METHOD PRIVATE Teach_OutOfTolerance_IsRejected
VAR_INST
    bRan : BOOL;
END_VAR
VAR
    stPlace : ST_SlotAddr := (nSide := 1, nColumn := 3, nLevel := 2);
END_VAR
TEST('Teach_OutOfTolerance_IsRejected');
IF bRan THEN
    TEST_FINISHED();
    RETURN;
END_IF
bRan := TRUE;

AssertFalse(Condition := fbRackReject.Teach(stPlace, fbRackReject.NominalX(stPlace) + 0.035, fbRackReject.NominalY(stPlace)),
            Message := '35 mm off the drawing means check the rack, not learn it');
AssertEquals_LREAL(Expected := fbRackReject.NominalX(stPlace), Actual := fbRackReject.TargetX(stPlace), Delta := 1.0E-9,
                   Message := 'a rejected teach must not change the target');

TEST_FINISHED();
END_METHOD

METHOD PRIVATE PutTake_BooksThePalletInAndOut
VAR_INST
    bRan : BOOL;
END_VAR
VAR
    stPlace : ST_SlotAddr := (nSide := 1, nColumn := 1, nLevel := 1);
END_VAR
TEST('PutTake_BooksThePalletInAndOut');
IF bRan THEN
    TEST_FINISHED();
    RETURN;
END_IF
bRan := TRUE;

AssertTrue(Condition := fbRackBook.Put(stPlace, 'LE0001'), Message := 'empty place must accept a pallet');
AssertTrue(Condition := fbRackBook.IsOccupied(stPlace), Message := 'place must be occupied after Put');
AssertEquals_STRING(Expected := 'LE0001', Actual := fbRackBook.LeIdAt(stPlace), Message := 'place must know its load unit');
AssertEquals_STRING(Expected := 'LE0001', Actual := fbRackBook.Take(stPlace), Message := 'Take must return the load unit');
AssertFalse(Condition := fbRackBook.IsOccupied(stPlace), Message := 'place must be free after Take');

TEST_FINISHED();
END_METHOD

METHOD PRIVATE Put_OnOccupiedPlace_IsRefused
VAR_INST
    bRan : BOOL;
END_VAR
VAR
    stPlace : ST_SlotAddr := (nSide := 2, nColumn := 7, nLevel := 4);
END_VAR
TEST('Put_OnOccupiedPlace_IsRefused');
IF bRan THEN
    TEST_FINISHED();
    RETURN;
END_IF
bRan := TRUE;

fbRackTwice.Put(stPlace, 'LE0001');
AssertFalse(Condition := fbRackTwice.Put(stPlace, 'LE0002'), Message := 'two pallets must never be booked into one place');
AssertEquals_STRING(Expected := 'LE0001', Actual := fbRackTwice.LeIdAt(stPlace), Message := 'first pallet must stay booked');

TEST_FINISHED();
END_METHOD

METHOD PRIVATE InvalidAddress_IsRejectedEverywhere
VAR_INST
    bRan : BOOL;
END_VAR
VAR
    stSide3 : ST_SlotAddr := (nSide := 3, nColumn := 1, nLevel := 1);
    stCol21 : ST_SlotAddr := (nSide := 1, nColumn := 21, nLevel := 1);
    stStationLevel2 : ST_SlotAddr := (nSide := 1, nColumn := 0, nLevel := 2);
END_VAR
TEST('InvalidAddress_IsRejectedEverywhere');
IF bRan THEN
    TEST_FINISHED();
    RETURN;
END_IF
bRan := TRUE;

AssertFalse(Condition := fbRackBad.IsValid(stSide3), Message := 'side 3 does not exist');
AssertFalse(Condition := fbRackBad.IsValid(stCol21), Message := 'column 21 does not exist');
AssertFalse(Condition := fbRackBad.IsValid(stStationLevel2), Message := 'the station has only level 1');
AssertFalse(Condition := fbRackBad.Put(stCol21, 'LE0001'), Message := 'no booking into an invalid address');

TEST_FINISHED();
END_METHOD

METHOD PRIVATE FindFree_SkipsOccupiedPlaces
VAR_INST
    bRan : BOOL;
END_VAR
VAR
    stA : ST_SlotAddr := (nSide := 1, nColumn := 1, nLevel := 1);
    stB : ST_SlotAddr := (nSide := 2, nColumn := 1, nLevel := 1);
    stFound : ST_SlotAddr;
END_VAR
TEST('FindFree_SkipsOccupiedPlaces');
IF bRan THEN
    TEST_FINISHED();
    RETURN;
END_IF
bRan := TRUE;

fbRackFree.Put(stA, 'LE0001');
fbRackFree.Put(stB, 'LE0002');
AssertTrue(Condition := fbRackFree.FindFree(stFound), Message := 'an almost empty rack has free places');
AssertEquals_INT(Expected := 1, Actual := stFound.nColumn, Message := 'nearest column first');
AssertEquals_INT(Expected := 2, Actual := stFound.nLevel, Message := 'level 1 is full on both sides -> level 2');

TEST_FINISHED();
END_METHOD

END_FUNCTION_BLOCK

// ---- Test/FB_Axis_Test.TcPOU
// Tests for FB_Axis, the simulated positioning axis. Each test drives the axis
// to the end inside one PLC cycle (simulated time), so they are fast.
FUNCTION_BLOCK FB_Axis_Test EXTENDS TcUnit.FB_TestSuite
VAR
    fbAxArrive  : FB_Axis(ipParent := 0, sNodeName := 'AxArrive');
    fbAxLong    : FB_Axis(ipParent := 0, sNodeName := 'AxLong');
    fbAxShort   : FB_Axis(ipParent := 0, sNodeName := 'AxShort');
    fbAxFault   : FB_Axis(ipParent := 0, sNodeName := 'AxFault');
    fbAxReset   : FB_Axis(ipParent := 0, sNodeName := 'AxReset');
END_VAR

Move_ArrivesInsideTheTolerance();
LongMove_TakesTheTrapezoidTime();
ShortMove_TakesTheTriangleTime();
DriveFault_WhileMoving_FailsTheMove();
Reset_AfterFault_AllowsTheNextMove();

METHOD PRIVATE Move_ArrivesInsideTheTolerance
VAR_INST
    bRan : BOOL;
END_VAR
VAR
    eResult : E_CmdResult;
    n : DINT;
END_VAR
TEST('Move_ArrivesInsideTheTolerance');
IF bRan THEN
    TEST_FINISHED();
    RETURN;
END_IF
bRan := TRUE;

FOR n := 1 TO 20000 DO
    eResult := fbAxArrive.MoveAbs(10.0);
    IF eResult <> E_CmdResult.eBusy THEN EXIT; END_IF
    fbAxArrive.Cyclic();
END_FOR
AssertTrue(Condition := eResult = E_CmdResult.eDone, Message := 'move must finish with eDone');
AssertEquals_LREAL(Expected := 10.0, Actual := fbAxArrive.lrActPos, Delta := fbAxArrive.lrTolerance, Message := 'axis must stand inside the tolerance');
AssertEquals_LREAL(Expected := 0.0, Actual := fbAxArrive.lrActVelo, Delta := 1.0E-9, Message := 'axis must stand still');

TEST_FINISHED();
END_METHOD

METHOD PRIVATE LongMove_TakesTheTrapezoidTime
VAR_INST
    bRan : BOOL;
END_VAR
VAR
    eResult : E_CmdResult;
    n : DINT;
    lrTime : LREAL;
END_VAR
TEST('LongMove_TakesTheTrapezoidTime');
IF bRan THEN
    TEST_FINISHED();
    RETURN;
END_IF
bRan := TRUE;

fbAxLong.lrVelocity := 3.0;
fbAxLong.lrAccel    := 0.6;
FOR n := 1 TO 20000 DO
    eResult := fbAxLong.MoveAbs(20.0);
    IF eResult <> E_CmdResult.eBusy THEN EXIT; END_IF
    fbAxLong.Cyclic();
    lrTime := lrTime + fbAxLong.lrCycleTime;
END_FOR
// 20 m >= v^2/a = 15 m -> top speed reached: t = s/v + v/a = 6.67 + 5.0 s
AssertEquals_LREAL(Expected := F_TravelTime(20.0, 3.0, 0.6), Actual := lrTime, Delta := 0.1, Message := 'move time must match s/v + v/a');

TEST_FINISHED();
END_METHOD

METHOD PRIVATE ShortMove_TakesTheTriangleTime
VAR_INST
    bRan : BOOL;
END_VAR
VAR
    eResult : E_CmdResult;
    n : DINT;
    lrTime : LREAL;
END_VAR
TEST('ShortMove_TakesTheTriangleTime');
IF bRan THEN
    TEST_FINISHED();
    RETURN;
END_IF
bRan := TRUE;

fbAxShort.lrVelocity := 3.0;
fbAxShort.lrAccel    := 0.6;
FOR n := 1 TO 20000 DO
    eResult := fbAxShort.MoveAbs(1.0);
    IF eResult <> E_CmdResult.eBusy THEN EXIT; END_IF
    fbAxShort.Cyclic();
    lrTime := lrTime + fbAxShort.lrCycleTime;
END_FOR
// 1 m < 15 m -> never reaches 3 m/s: t = 2 * sqrt(s/a) = 2.58 s
AssertEquals_LREAL(Expected := F_TravelTime(1.0, 3.0, 0.6), Actual := lrTime, Delta := 0.1, Message := 'short move must follow the triangle profile');

TEST_FINISHED();
END_METHOD

METHOD PRIVATE DriveFault_WhileMoving_FailsTheMove
VAR_INST
    bRan : BOOL;
END_VAR
VAR
    eResult : E_CmdResult;
    n : DINT;
END_VAR
TEST('DriveFault_WhileMoving_FailsTheMove');
IF bRan THEN
    TEST_FINISHED();
    RETURN;
END_IF
bRan := TRUE;

FOR n := 1 TO 50 DO
    fbAxFault.MoveAbs(5.0);
    fbAxFault.Cyclic();
END_FOR
fbAxFault.bDriveFault := TRUE;
fbAxFault.Cyclic();
eResult := fbAxFault.MoveAbs(5.0);
AssertTrue(Condition := eResult = E_CmdResult.eError, Message := 'a drive fault during a move must give eError');
AssertEquals_LREAL(Expected := 0.0, Actual := fbAxFault.lrActVelo, Delta := 1.0E-9, Message := 'a faulted axis must stand still');

TEST_FINISHED();
END_METHOD

METHOD PRIVATE Reset_AfterFault_AllowsTheNextMove
VAR_INST
    bRan : BOOL;
END_VAR
VAR
    eResult : E_CmdResult;
    n : DINT;
END_VAR
TEST('Reset_AfterFault_AllowsTheNextMove');
IF bRan THEN
    TEST_FINISHED();
    RETURN;
END_IF
bRan := TRUE;

fbAxReset.MoveAbs(5.0);
fbAxReset.Cyclic();
fbAxReset.bDriveFault := TRUE;
fbAxReset.Cyclic();
fbAxReset.bDriveFault := FALSE;
fbAxReset.Reset();
FOR n := 1 TO 20000 DO
    eResult := fbAxReset.MoveAbs(2.0);
    IF eResult <> E_CmdResult.eBusy THEN EXIT; END_IF
    fbAxReset.Cyclic();
END_FOR
AssertTrue(Condition := eResult = E_CmdResult.eDone, Message := 'after Reset a new move must work');

TEST_FINISHED();
END_METHOD

END_FUNCTION_BLOCK

// ---- Performance/F_TravelTime.TcPOU
// Time for one axis to travel lrDist with a trapezoid profile [s]:
// reaches top speed if lrDist >= v^2/a, otherwise a triangle profile.
FUNCTION F_TravelTime : LREAL
VAR_INPUT
    lrDist  : LREAL;   // [m]
    lrVelo  : LREAL;   // max. speed [m/s]
    lrAccel : LREAL;   // acceleration = deceleration [m/s2]
END_VAR
VAR
    lrD : LREAL;
END_VAR

lrD := ABS(lrDist);
IF lrD <= 0.0 OR lrVelo <= 0.0 OR lrAccel <= 0.0 THEN
    F_TravelTime := 0.0;
ELSIF lrD >= lrVelo * lrVelo / lrAccel THEN
    F_TravelTime := lrD / lrVelo + lrVelo / lrAccel;
ELSE
    F_TravelTime := 2.0 * SQRT(lrD / lrAccel);
END_IF

END_FUNCTION

// ---- Test/FB_ConveyorZone_Test.TcPOU
// Tests for FB_ConveyorZone, the standard conveyor block of the pre-zone.
FUNCTION_BLOCK FB_ConveyorZone_Test EXTENDS TcUnit.FB_TestSuite
VAR
    fbZoneIn    : FB_ConveyorZone(ipParent := 0, sNodeName := 'ZoneIn');
    fbZoneFull  : FB_ConveyorZone(ipParent := 0, sNodeName := 'ZoneFull');
    fbZoneOut   : FB_ConveyorZone(ipParent := 0, sNodeName := 'ZoneOut');
    fbZoneJam   : FB_ConveyorZone(ipParent := 0, sNodeName := 'ZoneJam');
END_VAR

Accept_RunsThePalletToTheEndLightBarrier();
Accept_OnOccupiedZone_IsRefused();
Deliver_EmptiesTheZoneWhenThePalletHasLeft();
LightBarrierNeverReached_IsAJam();

METHOD PRIVATE Accept_RunsThePalletToTheEndLightBarrier
VAR_INST
    bRan : BOOL;
END_VAR
VAR
    n : DINT;
    lrTime : LREAL;
END_VAR
TEST('Accept_RunsThePalletToTheEndLightBarrier');
IF bRan THEN
    TEST_FINISHED();
    RETURN;
END_IF
bRan := TRUE;

AssertTrue(Condition := fbZoneIn.Accept('LE0001'), Message := 'an empty zone must accept a pallet');
FOR n := 1 TO 5000 DO
    fbZoneIn.Cyclic();
    lrTime := lrTime + fbZoneIn.lrCycleTime;
    IF fbZoneIn.eState = E_ZoneState.eOccupied THEN EXIT; END_IF
END_FOR
AssertTrue(Condition := fbZoneIn.eState = E_ZoneState.eOccupied, Message := 'pallet must stop at the end light barrier');
AssertFalse(Condition := fbZoneIn.bMotorOn, Message := 'motor must be off when the pallet has arrived');
AssertEquals_LREAL(Expected := 8.0, Actual := lrTime, Delta := 0.05, Message := '1.6 m at 0.2 m/s = 8 s');
AssertEquals_STRING(Expected := 'LE0001', Actual := fbZoneIn.sLeId, Message := 'zone must know its pallet');

TEST_FINISHED();
END_METHOD

METHOD PRIVATE Accept_OnOccupiedZone_IsRefused
VAR_INST
    bRan : BOOL;
END_VAR
VAR
    n : DINT;
END_VAR
TEST('Accept_OnOccupiedZone_IsRefused');
IF bRan THEN
    TEST_FINISHED();
    RETURN;
END_IF
bRan := TRUE;

fbZoneFull.Accept('LE0001');
FOR n := 1 TO 5000 DO
    fbZoneFull.Cyclic();
END_FOR
AssertFalse(Condition := fbZoneFull.Accept('LE0002'), Message := 'a zone holds one pallet only');

TEST_FINISHED();
END_METHOD

METHOD PRIVATE Deliver_EmptiesTheZoneWhenThePalletHasLeft
VAR_INST
    bRan : BOOL;
END_VAR
VAR
    n : DINT;
    eResult : E_CmdResult;
END_VAR
TEST('Deliver_EmptiesTheZoneWhenThePalletHasLeft');
IF bRan THEN
    TEST_FINISHED();
    RETURN;
END_IF
bRan := TRUE;

fbZoneOut.Accept('LE0001');
FOR n := 1 TO 5000 DO
    fbZoneOut.Cyclic();
END_FOR
FOR n := 1 TO 5000 DO
    eResult := fbZoneOut.Deliver();
    IF eResult <> E_CmdResult.eBusy THEN EXIT; END_IF
    fbZoneOut.Cyclic();
END_FOR
AssertTrue(Condition := eResult = E_CmdResult.eDone, Message := 'deliver must end with eDone');
AssertTrue(Condition := fbZoneOut.eState = E_ZoneState.eEmpty, Message := 'zone must be empty after delivering');
AssertEquals_STRING(Expected := '', Actual := fbZoneOut.sLeId, Message := 'zone must forget the pallet');

TEST_FINISHED();
END_METHOD

METHOD PRIVATE LightBarrierNeverReached_IsAJam
VAR_INST
    bRan : BOOL;
END_VAR
VAR
    n : DINT;
END_VAR
TEST('LightBarrierNeverReached_IsAJam');
IF bRan THEN
    TEST_FINISHED();
    RETURN;
END_IF
bRan := TRUE;

fbZoneJam.bSimulate    := FALSE;   // real sensor that never switches
fbZoneJam.lrJamTimeout := 5.0;
fbZoneJam.Accept('LE0001');
FOR n := 1 TO 600 DO
    fbZoneJam.Cyclic();
END_FOR
AssertTrue(Condition := fbZoneJam.eState = E_ZoneState.eFault, Message := 'no light barrier after the jam time must be a fault');
AssertFalse(Condition := fbZoneJam.bMotorOn, Message := 'motor must stop on a jam');

TEST_FINISHED();
END_METHOD

END_FUNCTION_BLOCK

// ---- Test/FB_IPoint_Test.TcPOU
// Tests for FB_IPoint, the contour check and barcode read before storage.
FUNCTION_BLOCK FB_IPoint_Test EXTENDS TcUnit.FB_TestSuite
VAR
    fbIpOk      : FB_IPoint;
    fbIpContour : FB_IPoint;
    fbIpNoRead  : FB_IPoint;
END_VAR

GoodPallet_IsOk();
Overhang_IsContourNio();
NoBarcode_IsNoReadNio();

METHOD PRIVATE GoodPallet_IsOk
VAR_INST
    bRan : BOOL;
END_VAR
TEST('GoodPallet_IsOk');
IF bRan THEN
    TEST_FINISHED();
    RETURN;
END_IF
bRan := TRUE;

fbIpOk.sBarcode := 'LE0001';
AssertTrue(Condition := fbIpOk.Check() = E_IPointResult.eOk, Message := 'clean contour and a read barcode = OK');

TEST_FINISHED();
END_METHOD

METHOD PRIVATE Overhang_IsContourNio
VAR_INST
    bRan : BOOL;
END_VAR
TEST('Overhang_IsContourNio');
IF bRan THEN
    TEST_FINISHED();
    RETURN;
END_IF
bRan := TRUE;

fbIpContour.sBarcode      := 'LE0001';
fbIpContour.bOverhangLeft := TRUE;
AssertTrue(Condition := fbIpContour.Check() = E_IPointResult.eNioContour, Message := 'overhang must be rejected');
AssertEquals_DINT(Expected := 1, Actual := fbIpContour.nNio, Message := 'NIO counter');

TEST_FINISHED();
END_METHOD

METHOD PRIVATE NoBarcode_IsNoReadNio
VAR_INST
    bRan : BOOL;
END_VAR
TEST('NoBarcode_IsNoReadNio');
IF bRan THEN
    TEST_FINISHED();
    RETURN;
END_IF
bRan := TRUE;

AssertTrue(Condition := fbIpNoRead.Check() = E_IPointResult.eNioNoRead, Message := 'no barcode must be rejected');

TEST_FINISHED();
END_METHOD

END_FUNCTION_BLOCK

// ---- Test/FB_MfrInterface_Test.TcPOU
// Tests for the telegram interface to the material flow computer: these are
// the interface test cases of the commissioning (Schnittstellentest).
FUNCTION_BLOCK FB_MfrInterface_Test EXTENDS TcUnit.FB_TestSuite
VAR
    fbRackOk : FB_Rack;
    fbSrmOk  : FB_Srm(ipParent := 0, sNodeName := 'SrmOk');
    fbMfrOk  : FB_MfrInterface;
    fbRackSeq : FB_Rack;
    fbSrmSeq  : FB_Srm(ipParent := 0, sNodeName := 'SrmSeq');
    fbMfrSeq  : FB_MfrInterface;
    fbRackDup : FB_Rack;
    fbSrmDup  : FB_Srm(ipParent := 0, sNodeName := 'SrmDup');
    fbMfrDup  : FB_MfrInterface;
    fbRackOcc : FB_Rack;
    fbSrmOcc  : FB_Srm(ipParent := 0, sNodeName := 'SrmOcc');
    fbMfrOcc  : FB_MfrInterface;
    fbRackEmpty : FB_Rack;
    fbSrmEmpty  : FB_Srm(ipParent := 0, sNodeName := 'SrmEmpty');
    fbMfrEmpty  : FB_MfrInterface;
    fbRackLe : FB_Rack;
    fbSrmLe  : FB_Srm(ipParent := 0, sNodeName := 'SrmLe');
    fbMfrLe  : FB_MfrInterface;
    fbRackAddr : FB_Rack;
    fbSrmAddr  : FB_Srm(ipParent := 0, sNodeName := 'SrmAddr');
    fbMfrAddr  : FB_MfrInterface;
    fbRackBusy : FB_Rack;
    fbSrmBusy  : FB_Srm(ipParent := 0, sNodeName := 'SrmBusy');
    fbMfrBusy  : FB_MfrInterface;
    fbRackDone : FB_Rack;
    fbSrmDone  : FB_Srm(ipParent := 0, sNodeName := 'SrmDone');
    fbMfrDone  : FB_MfrInterface;
    fbRackAck : FB_Rack;
    fbSrmAck  : FB_Srm(ipParent := 0, sNodeName := 'SrmAck');
    fbMfrAck  : FB_MfrInterface;
END_VAR

ValidOrder_IsAcknowledgedAndStarted();
WrongSequenceNumber_IsRejected();
DuplicateOrder_IsRejected();
TargetOccupied_IsRejected();
SourceEmpty_IsRejected();
WrongLoadUnit_IsRejected();
InvalidAddress_IsRejected();
SecondOrderWhileBusy_IsRejected();
FinishedJob_SendsTdon_AndMissingAckTimesOut();
Tack_ClearsTheWaitForAcknowledge();

METHOD PRIVATE ValidOrder_IsAcknowledgedAndStarted
VAR_INST
    bRan : BOOL;
END_VAR
VAR
    stTel, stAns : ST_Telegram;
    stStation : ST_SlotAddr := (nSide := 1, nColumn := 0, nLevel := 1);
    stPlace : ST_SlotAddr := (nSide := 1, nColumn := 2, nLevel := 1);
    stOther : ST_SlotAddr := (nSide := 2, nColumn := 6, nLevel := 3);
    stBad   : ST_SlotAddr := (nSide := 1, nColumn := 30, nLevel := 1);
    n : DINT;
END_VAR
TEST('ValidOrder_IsAcknowledgedAndStarted');
IF bRan THEN
    TEST_FINISHED();
    RETURN;
END_IF
bRan := TRUE;

fbMfrOk.Init(fbRackOk, fbSrmOk);
fbSrmOk.Init(fbRackOk);
fbRackOk.Put(stStation, 'LE0001');
stTel.sType := 'TORD'; stTel.nSeq := 1; stTel.nOrder := 1; stTel.sLeId := 'LE0001';
stTel.stSource := stStation; stTel.stTarget := stPlace;
stAns := fbMfrOk.Receive(stTel);
AssertEquals_STRING(Expected := 'TACK', Actual := stAns.sType, Message := 'a valid order must be acknowledged');
AssertEquals_INT(Expected := GVL_Mfr.cStatusOk, Actual := stAns.nStatus, Message := 'status OK');
AssertEquals_DINT(Expected := 1, Actual := fbMfrOk.ActiveOrder, Message := 'order must be active');

TEST_FINISHED();
END_METHOD

METHOD PRIVATE WrongSequenceNumber_IsRejected
VAR_INST
    bRan : BOOL;
END_VAR
VAR
    stTel, stAns : ST_Telegram;
    stStation : ST_SlotAddr := (nSide := 1, nColumn := 0, nLevel := 1);
    stPlace : ST_SlotAddr := (nSide := 1, nColumn := 2, nLevel := 1);
    stOther : ST_SlotAddr := (nSide := 2, nColumn := 6, nLevel := 3);
    stBad   : ST_SlotAddr := (nSide := 1, nColumn := 30, nLevel := 1);
    n : DINT;
END_VAR
TEST('WrongSequenceNumber_IsRejected');
IF bRan THEN
    TEST_FINISHED();
    RETURN;
END_IF
bRan := TRUE;

fbMfrSeq.Init(fbRackSeq, fbSrmSeq);
fbSrmSeq.Init(fbRackSeq);
fbRackSeq.Put(stStation, 'LE0001');
stTel.sType := 'TORD'; stTel.nSeq := 2; stTel.nOrder := 1; stTel.sLeId := 'LE0001';
stTel.stSource := stStation; stTel.stTarget := stPlace;
stAns := fbMfrSeq.Receive(stTel);
AssertEquals_INT(Expected := GVL_Mfr.cWrongSequence, Actual := stAns.nStatus, Message := 'first telegram must carry seq 1');
AssertEquals_DINT(Expected := 0, Actual := fbMfrSeq.ActiveOrder, Message := 'nothing may start');

TEST_FINISHED();
END_METHOD

METHOD PRIVATE DuplicateOrder_IsRejected
VAR_INST
    bRan : BOOL;
END_VAR
VAR
    stTel, stAns : ST_Telegram;
    stStation : ST_SlotAddr := (nSide := 1, nColumn := 0, nLevel := 1);
    stPlace : ST_SlotAddr := (nSide := 1, nColumn := 2, nLevel := 1);
    stOther : ST_SlotAddr := (nSide := 2, nColumn := 6, nLevel := 3);
    stBad   : ST_SlotAddr := (nSide := 1, nColumn := 30, nLevel := 1);
    n : DINT;
END_VAR
TEST('DuplicateOrder_IsRejected');
IF bRan THEN
    TEST_FINISHED();
    RETURN;
END_IF
bRan := TRUE;

fbMfrDup.Init(fbRackDup, fbSrmDup);
fbSrmDup.Init(fbRackDup);
fbRackDup.Put(stStation, 'LE0001');
stTel.sType := 'TORD'; stTel.nSeq := 1; stTel.nOrder := 7; stTel.sLeId := 'LE0001';
stTel.stSource := stStation; stTel.stTarget := stPlace;
fbMfrDup.Receive(stTel);
stTel.nSeq := 2;
stAns := fbMfrDup.Receive(stTel);
AssertEquals_INT(Expected := GVL_Mfr.cDuplicateOrder, Actual := stAns.nStatus, Message := 'same order number twice must be rejected');

TEST_FINISHED();
END_METHOD

METHOD PRIVATE TargetOccupied_IsRejected
VAR_INST
    bRan : BOOL;
END_VAR
VAR
    stTel, stAns : ST_Telegram;
    stStation : ST_SlotAddr := (nSide := 1, nColumn := 0, nLevel := 1);
    stPlace : ST_SlotAddr := (nSide := 1, nColumn := 2, nLevel := 1);
    stOther : ST_SlotAddr := (nSide := 2, nColumn := 6, nLevel := 3);
    stBad   : ST_SlotAddr := (nSide := 1, nColumn := 30, nLevel := 1);
    n : DINT;
END_VAR
TEST('TargetOccupied_IsRejected');
IF bRan THEN
    TEST_FINISHED();
    RETURN;
END_IF
bRan := TRUE;

fbMfrOcc.Init(fbRackOcc, fbSrmOcc);
fbSrmOcc.Init(fbRackOcc);
fbRackOcc.Put(stStation, 'LE0001');fbRackOcc.Put(stPlace, 'LE0099');
stTel.sType := 'TORD'; stTel.nSeq := 1; stTel.nOrder := 1; stTel.sLeId := 'LE0001';
stTel.stSource := stStation; stTel.stTarget := stPlace;
stAns := fbMfrOcc.Receive(stTel);
AssertEquals_INT(Expected := GVL_Mfr.cSlotOccupied, Actual := stAns.nStatus, Message := 'never store into an occupied place');

TEST_FINISHED();
END_METHOD

METHOD PRIVATE SourceEmpty_IsRejected
VAR_INST
    bRan : BOOL;
END_VAR
VAR
    stTel, stAns : ST_Telegram;
    stStation : ST_SlotAddr := (nSide := 1, nColumn := 0, nLevel := 1);
    stPlace : ST_SlotAddr := (nSide := 1, nColumn := 2, nLevel := 1);
    stOther : ST_SlotAddr := (nSide := 2, nColumn := 6, nLevel := 3);
    stBad   : ST_SlotAddr := (nSide := 1, nColumn := 30, nLevel := 1);
    n : DINT;
END_VAR
TEST('SourceEmpty_IsRejected');
IF bRan THEN
    TEST_FINISHED();
    RETURN;
END_IF
bRan := TRUE;

fbMfrEmpty.Init(fbRackEmpty, fbSrmEmpty);
fbSrmEmpty.Init(fbRackEmpty);
fbRackEmpty.Put(stStation, 'LE0001');
stTel.sType := 'TORD'; stTel.nSeq := 1; stTel.nOrder := 1; stTel.sLeId := 'LE0005';
stTel.stSource := stOther; stTel.stTarget := stPlace;
stAns := fbMfrEmpty.Receive(stTel);
AssertEquals_INT(Expected := GVL_Mfr.cSlotEmpty, Actual := stAns.nStatus, Message := 'no pick from an empty place');

TEST_FINISHED();
END_METHOD

METHOD PRIVATE WrongLoadUnit_IsRejected
VAR_INST
    bRan : BOOL;
END_VAR
VAR
    stTel, stAns : ST_Telegram;
    stStation : ST_SlotAddr := (nSide := 1, nColumn := 0, nLevel := 1);
    stPlace : ST_SlotAddr := (nSide := 1, nColumn := 2, nLevel := 1);
    stOther : ST_SlotAddr := (nSide := 2, nColumn := 6, nLevel := 3);
    stBad   : ST_SlotAddr := (nSide := 1, nColumn := 30, nLevel := 1);
    n : DINT;
END_VAR
TEST('WrongLoadUnit_IsRejected');
IF bRan THEN
    TEST_FINISHED();
    RETURN;
END_IF
bRan := TRUE;

fbMfrLe.Init(fbRackLe, fbSrmLe);
fbSrmLe.Init(fbRackLe);
fbRackLe.Put(stStation, 'LE0001');
stTel.sType := 'TORD'; stTel.nSeq := 1; stTel.nOrder := 1; stTel.sLeId := 'LE0042';
stTel.stSource := stStation; stTel.stTarget := stPlace;
stAns := fbMfrLe.Receive(stTel);
AssertEquals_INT(Expected := GVL_Mfr.cLeMismatch, Actual := stAns.nStatus, Message := 'ordered pallet must be the one at the source');

TEST_FINISHED();
END_METHOD

METHOD PRIVATE InvalidAddress_IsRejected
VAR_INST
    bRan : BOOL;
END_VAR
VAR
    stTel, stAns : ST_Telegram;
    stStation : ST_SlotAddr := (nSide := 1, nColumn := 0, nLevel := 1);
    stPlace : ST_SlotAddr := (nSide := 1, nColumn := 2, nLevel := 1);
    stOther : ST_SlotAddr := (nSide := 2, nColumn := 6, nLevel := 3);
    stBad   : ST_SlotAddr := (nSide := 1, nColumn := 30, nLevel := 1);
    n : DINT;
END_VAR
TEST('InvalidAddress_IsRejected');
IF bRan THEN
    TEST_FINISHED();
    RETURN;
END_IF
bRan := TRUE;

fbMfrAddr.Init(fbRackAddr, fbSrmAddr);
fbSrmAddr.Init(fbRackAddr);
fbRackAddr.Put(stStation, 'LE0001');
stTel.sType := 'TORD'; stTel.nSeq := 1; stTel.nOrder := 1; stTel.sLeId := 'LE0001';
stTel.stSource := stStation; stTel.stTarget := stBad;
stAns := fbMfrAddr.Receive(stTel);
AssertEquals_INT(Expected := GVL_Mfr.cInvalidAddress, Actual := stAns.nStatus, Message := 'column 30 does not exist');

TEST_FINISHED();
END_METHOD

METHOD PRIVATE SecondOrderWhileBusy_IsRejected
VAR_INST
    bRan : BOOL;
END_VAR
VAR
    stTel, stAns : ST_Telegram;
    stStation : ST_SlotAddr := (nSide := 1, nColumn := 0, nLevel := 1);
    stPlace : ST_SlotAddr := (nSide := 1, nColumn := 2, nLevel := 1);
    stOther : ST_SlotAddr := (nSide := 2, nColumn := 6, nLevel := 3);
    stBad   : ST_SlotAddr := (nSide := 1, nColumn := 30, nLevel := 1);
    n : DINT;
END_VAR
TEST('SecondOrderWhileBusy_IsRejected');
IF bRan THEN
    TEST_FINISHED();
    RETURN;
END_IF
bRan := TRUE;

fbMfrBusy.Init(fbRackBusy, fbSrmBusy);
fbSrmBusy.Init(fbRackBusy);
fbRackBusy.Put(stStation, 'LE0001');
stTel.sType := 'TORD'; stTel.nSeq := 1; stTel.nOrder := 1; stTel.sLeId := 'LE0001';
stTel.stSource := stStation; stTel.stTarget := stPlace;
fbMfrBusy.Receive(stTel);
fbRackBusy.Put(stOther, 'LE0002');
stTel.nSeq := 2; stTel.nOrder := 2; stTel.sLeId := 'LE0002'; stTel.stSource := stOther;
stTel.stTarget := stPlace;
stTel.stTarget.nColumn := 9;   // free place (1,9,1)
stAns := fbMfrBusy.Receive(stTel);
AssertEquals_INT(Expected := GVL_Mfr.cSrmBusy, Actual := stAns.nStatus, Message := 'one order at a time');

TEST_FINISHED();
END_METHOD

METHOD PRIVATE FinishedJob_SendsTdon_AndMissingAckTimesOut
VAR_INST
    bRan : BOOL;
END_VAR
VAR
    stTel, stAns : ST_Telegram;
    stStation : ST_SlotAddr := (nSide := 1, nColumn := 0, nLevel := 1);
    stPlace : ST_SlotAddr := (nSide := 1, nColumn := 2, nLevel := 1);
    stOther : ST_SlotAddr := (nSide := 2, nColumn := 6, nLevel := 3);
    stBad   : ST_SlotAddr := (nSide := 1, nColumn := 30, nLevel := 1);
    n : DINT;
END_VAR
TEST('FinishedJob_SendsTdon_AndMissingAckTimesOut');
IF bRan THEN
    TEST_FINISHED();
    RETURN;
END_IF
bRan := TRUE;

fbMfrDone.Init(fbRackDone, fbSrmDone);
fbSrmDone.Init(fbRackDone);
fbRackDone.Put(stStation, 'LE0001');
stTel.sType := 'TORD'; stTel.nSeq := 1; stTel.nOrder := 1; stTel.sLeId := 'LE0001';
stTel.stSource := stStation; stTel.stTarget := stPlace;
fbSrmDone.SetMode(E_OpMode.eAutomatic);
fbMfrDone.Receive(stTel);
FOR n := 1 TO 30000 DO
    fbSrmDone.Cyclic();
    fbMfrDone.Cyclic();
    IF fbMfrDone.nOutboxCount > 0 THEN EXIT; END_IF
END_FOR
AssertEquals_STRING(Expected := 'TDON', Actual := fbMfrDone.stOutbox.sType, Message := 'finished order must be reported with TDON');
AssertEquals_DINT(Expected := 1, Actual := fbMfrDone.stOutbox.nOrder, Message := 'TDON must carry the order number');
FOR n := 1 TO 600 DO   // 6 s without TACK
    fbMfrDone.Cyclic();
END_FOR
AssertTrue(Condition := fbMfrDone.bAckTimeout, Message := 'missing TACK must time out');
AssertEquals_INT(Expected := GVL_Mfr.cAckTimeout, Actual := fbMfrDone.nLastStatus, Message := 'status 30');

TEST_FINISHED();
END_METHOD

METHOD PRIVATE Tack_ClearsTheWaitForAcknowledge
VAR_INST
    bRan : BOOL;
END_VAR
VAR
    stTel, stAns : ST_Telegram;
    stStation : ST_SlotAddr := (nSide := 1, nColumn := 0, nLevel := 1);
    stPlace : ST_SlotAddr := (nSide := 1, nColumn := 2, nLevel := 1);
    stOther : ST_SlotAddr := (nSide := 2, nColumn := 6, nLevel := 3);
    stBad   : ST_SlotAddr := (nSide := 1, nColumn := 30, nLevel := 1);
    n : DINT;
END_VAR
TEST('Tack_ClearsTheWaitForAcknowledge');
IF bRan THEN
    TEST_FINISHED();
    RETURN;
END_IF
bRan := TRUE;

fbMfrAck.Init(fbRackAck, fbSrmAck);
fbSrmAck.Init(fbRackAck);
fbRackAck.Put(stStation, 'LE0001');
stTel.sType := 'TORD'; stTel.nSeq := 1; stTel.nOrder := 1; stTel.sLeId := 'LE0001';
stTel.stSource := stStation; stTel.stTarget := stPlace;
fbSrmAck.SetMode(E_OpMode.eAutomatic);
fbMfrAck.Receive(stTel);
FOR n := 1 TO 30000 DO
    fbSrmAck.Cyclic();
    fbMfrAck.Cyclic();
    IF fbMfrAck.nOutboxCount > 0 THEN EXIT; END_IF
END_FOR
stTel.sType := 'TACK'; stTel.nSeq := 2; stTel.nOrder := 1;
fbMfrAck.Receive(stTel);
FOR n := 1 TO 600 DO
    fbMfrAck.Cyclic();
END_FOR
AssertFalse(Condition := fbMfrAck.AwaitingAck, Message := 'TACK must end the wait');
AssertFalse(Condition := fbMfrAck.bAckTimeout, Message := 'acknowledged TDON must not time out');

TEST_FINISHED();
END_METHOD

END_FUNCTION_BLOCK

// ---- Test/FB_Srm_Test.TcPOU
// Tests for FB_Srm, the storage and retrieval machine: whole jobs run in
// simulated time, and the double cycle is checked against FEM 9.851.
FUNCTION_BLOCK FB_Srm_Test EXTENDS TcUnit.FB_TestSuite
VAR
    fbRackStore : FB_Rack;
    fbSrmStore  : FB_Srm(ipParent := 0, sNodeName := 'SrmStore');
    fbRackGet : FB_Rack;
    fbSrmGet  : FB_Srm(ipParent := 0, sNodeName := 'SrmGet');
    fbRackOcc : FB_Rack;
    fbSrmOcc  : FB_Srm(ipParent := 0, sNodeName := 'SrmOcc');
    fbRackFault : FB_Rack;
    fbSrmFault  : FB_Srm(ipParent := 0, sNodeName := 'SrmFault');
    fbRackFem : FB_Rack;
    fbSrmFem  : FB_Srm(ipParent := 0, sNodeName := 'SrmFem');
END_VAR

StoreJob_MovesThePalletFromStationIntoThePlace();
RetrieveJob_BringsThePalletToTheStation();
StartJob_IntoOccupiedPlace_IsRefused();
TravelFault_StopsTheJobWithoutLosingThePallet();
DoubleCycle_MatchesTheFem9851Calculation();

METHOD PRIVATE StoreJob_MovesThePalletFromStationIntoThePlace
VAR_INST
    bRan : BOOL;
END_VAR
VAR
    stStation : ST_SlotAddr := (nSide := 1, nColumn := 0, nLevel := 1);
    stPlace : ST_SlotAddr := (nSide := 2, nColumn := 4, nLevel := 3);
    n : DINT;
END_VAR
TEST('StoreJob_MovesThePalletFromStationIntoThePlace');
IF bRan THEN
    TEST_FINISHED();
    RETURN;
END_IF
bRan := TRUE;

fbSrmStore.Init(fbRackStore);
fbSrmStore.SetMode(E_OpMode.eAutomatic);
fbRackStore.Put(stStation, 'LE0001');
AssertTrue(Condition := fbSrmStore.StartJob(stStation, stPlace), Message := 'job must be accepted');
FOR n := 1 TO 30000 DO
    fbSrmStore.Cyclic();
    IF fbSrmStore.bJobDone OR fbSrmStore.bFault THEN EXIT; END_IF
END_FOR
AssertTrue(Condition := fbSrmStore.bJobDone, Message := 'store job must finish');
AssertEquals_STRING(Expected := 'LE0001', Actual := fbRackStore.LeIdAt(stPlace), Message := 'pallet must be booked into the place');
AssertFalse(Condition := fbRackStore.IsOccupied(stStation), Message := 'station must be free');
AssertEquals_LREAL(Expected := fbRackStore.TargetX(stPlace), Actual := fbSrmStore.TravelPos, Delta := 0.002, Message := 'RBG must stand at the place');
AssertEquals_LREAL(Expected := 0.0, Actual := fbSrmStore.ForkActPos, Delta := 0.002, Message := 'fork must be back in the middle');

TEST_FINISHED();
END_METHOD

METHOD PRIVATE RetrieveJob_BringsThePalletToTheStation
VAR_INST
    bRan : BOOL;
END_VAR
VAR
    stStation : ST_SlotAddr := (nSide := 1, nColumn := 0, nLevel := 1);
    stPlace : ST_SlotAddr := (nSide := 2, nColumn := 4, nLevel := 3);
    n : DINT;
END_VAR
TEST('RetrieveJob_BringsThePalletToTheStation');
IF bRan THEN
    TEST_FINISHED();
    RETURN;
END_IF
bRan := TRUE;

fbSrmGet.Init(fbRackGet);
fbSrmGet.SetMode(E_OpMode.eAutomatic);
fbRackGet.Put(stPlace, 'LE0002');
fbSrmGet.StartJob(stPlace, stStation);
FOR n := 1 TO 30000 DO
    fbSrmGet.Cyclic();
    IF fbSrmGet.bJobDone OR fbSrmGet.bFault THEN EXIT; END_IF
END_FOR
AssertEquals_STRING(Expected := 'LE0002', Actual := fbRackGet.LeIdAt(stStation), Message := 'pallet must arrive at the station');

TEST_FINISHED();
END_METHOD

METHOD PRIVATE StartJob_IntoOccupiedPlace_IsRefused
VAR_INST
    bRan : BOOL;
END_VAR
VAR
    stStation : ST_SlotAddr := (nSide := 1, nColumn := 0, nLevel := 1);
    stPlace : ST_SlotAddr := (nSide := 2, nColumn := 4, nLevel := 3);
    n : DINT;
END_VAR
TEST('StartJob_IntoOccupiedPlace_IsRefused');
IF bRan THEN
    TEST_FINISHED();
    RETURN;
END_IF
bRan := TRUE;

fbSrmOcc.Init(fbRackOcc);
fbRackOcc.Put(stStation, 'LE0001');
fbRackOcc.Put(stPlace, 'LE0002');
AssertFalse(Condition := fbSrmOcc.StartJob(stStation, stPlace), Message := 'target occupied -> no job');

TEST_FINISHED();
END_METHOD

METHOD PRIVATE TravelFault_StopsTheJobWithoutLosingThePallet
VAR_INST
    bRan : BOOL;
END_VAR
VAR
    stStation : ST_SlotAddr := (nSide := 1, nColumn := 0, nLevel := 1);
    stPlace : ST_SlotAddr := (nSide := 2, nColumn := 4, nLevel := 3);
    n : DINT;
END_VAR
TEST('TravelFault_StopsTheJobWithoutLosingThePallet');
IF bRan THEN
    TEST_FINISHED();
    RETURN;
END_IF
bRan := TRUE;

fbSrmFault.Init(fbRackFault);
fbSrmFault.SetMode(E_OpMode.eAutomatic);
fbRackFault.Put(stPlace, 'LE0003');
fbSrmFault.StartJob(stPlace, stStation);
FOR n := 1 TO 100 DO
    fbSrmFault.Cyclic();
END_FOR
fbSrmFault.InjectTravelFault(TRUE);
FOR n := 1 TO 10 DO
    fbSrmFault.Cyclic();
END_FOR
AssertTrue(Condition := fbSrmFault.bFault, Message := 'a travel fault must stop the job');
AssertFalse(Condition := fbSrmFault.bJobDone, Message := 'faulted job is not done');
AssertEquals_STRING(Expected := 'LE0003', Actual := fbRackFault.LeIdAt(stPlace), Message := 'pallet must still be booked where it is');

TEST_FINISHED();
END_METHOD

METHOD PRIVATE DoubleCycle_MatchesTheFem9851Calculation
VAR_INST
    bRan : BOOL;
END_VAR
VAR
    stStation : ST_SlotAddr := (nSide := 1, nColumn := 0, nLevel := 1);
    stP1 : ST_SlotAddr := (nSide := 1, nColumn := 4, nLevel := 6);   // ~ (1/5 L, 2/3 H)
    stP2 : ST_SlotAddr := (nSide := 1, nColumn := 13, nLevel := 2);  // ~ (2/3 L, 1/5 H)
    stKin : ST_SrmKinematics := (lrVeloX := 3.0, lrAccelX := 0.6, lrVeloY := 1.5, lrAccelY := 0.8, lrVeloZ := 0.6, lrAccelZ := 0.6);
    n : DINT;
    lrMeasured, lrCalc : LREAL;
END_VAR
TEST('DoubleCycle_MatchesTheFem9851Calculation');
IF bRan THEN
    TEST_FINISHED();
    RETURN;
END_IF
bRan := TRUE;

fbSrmFem.Init(fbRackFem);
// 1. home to the station
fbSrmFem.SetMode(E_OpMode.eHoming);
FOR n := 1 TO 3000 DO
    fbSrmFem.Cyclic();
END_FOR
fbSrmFem.SetMode(E_OpMode.eAutomatic);
// 2. store at P1, then retrieve from P2 = one double cycle
fbRackFem.Put(stStation, 'LE0001');
fbRackFem.Put(stP2, 'LE0002');
fbSrmFem.StartJob(stStation, stP1);
FOR n := 1 TO 30000 DO
    fbSrmFem.Cyclic();
    IF fbSrmFem.bJobDone THEN EXIT; END_IF
END_FOR
lrMeasured := fbSrmFem.lrLastJobTime;
fbSrmFem.StartJob(stP2, stStation);
FOR n := 1 TO 30000 DO
    fbSrmFem.Cyclic();
    IF fbSrmFem.bJobDone THEN EXIT; END_IF
END_FOR
lrMeasured := lrMeasured + fbSrmFem.lrLastJobTime;

lrCalc := F_DoubleCycleTime(fbRackFem.NominalX(stP1), fbRackFem.NominalY(stP1) - GVL_Rack.cOffsetY,
                            fbRackFem.NominalX(stP2), fbRackFem.NominalY(stP2) - GVL_Rack.cOffsetY, stKin);
GVL_Test.lrDoubleCycleCalc     := lrCalc;
GVL_Test.lrDoubleCycleMeasured := lrMeasured;
IF lrMeasured > 0.0 THEN
    GVL_Test.lrDoubleCyclesPerHour := 3600.0 / lrMeasured;
END_IF
AssertEquals_LREAL(Expected := lrCalc, Actual := lrMeasured, Delta := 0.05 * lrCalc,
                   Message := 'simulated double cycle must be within 5 % of the FEM 9.851 calculation');

TEST_FINISHED();
END_METHOD

END_FUNCTION_BLOCK

// ---- Performance/F_DoubleCycleTime.TcPOU
// Double cycle as in the FEM 9.851 performance proof: from the transfer
// station store a pallet at P1, travel empty to P2, retrieve a pallet there and
// bring it back to the station. P1 and P2 are the reference places given as
// coordinates relative to the transfer station.
// FEM 9.851 places them at P1 = (1/5 L, 2/3 H) and P2 = (2/3 L, 1/5 H)
// (rack length L, rack height H) - see FB_Srm_Test.DoubleCycle_MatchesTheFem9851Calculation.
FUNCTION F_DoubleCycleTime : LREAL
VAR_INPUT
    lrX1, lrY1 : LREAL;   // P1 relative to the station [m]
    lrX2, lrY2 : LREAL;   // P2 relative to the station [m]
    stKin      : ST_SrmKinematics;
END_VAR

F_DoubleCycleTime := 4.0 * F_LoadHandlingTime(stKin)          // 2 x pick, 2 x deposit
                   + F_MoveTime(lrX1, lrY1, stKin)              // station -> P1 (loaded)
                   + F_MoveTime(lrX2 - lrX1, lrY2 - lrY1, stKin) // P1 -> P2 (empty)
                   + F_MoveTime(lrX2, lrY2, stKin);             // P2 -> station (loaded)

END_FUNCTION

// ---- Performance/F_LoadHandlingTime.TcPOU
// One pick or one deposit at a place: fork out, lift or lower, fork in.
FUNCTION F_LoadHandlingTime : LREAL
VAR_INPUT
    stKin : ST_SrmKinematics;
END_VAR

F_LoadHandlingTime := 2.0 * F_TravelTime(GVL_Rack.cForkStroke, stKin.lrVeloZ, stKin.lrAccelZ)
                    + F_TravelTime(GVL_Rack.cLiftStroke, stKin.lrVeloY, stKin.lrAccelY);

END_FUNCTION

// ---- Performance/F_MoveTime.TcPOU
// Travel and hoist run at the same time, so a move takes as long as the slower axis.
FUNCTION F_MoveTime : LREAL
VAR_INPUT
    lrDx  : LREAL;
    lrDy  : LREAL;
    stKin : ST_SrmKinematics;
END_VAR

F_MoveTime := MAX(F_TravelTime(lrDx, stKin.lrVeloX, stKin.lrAccelX),
                  F_TravelTime(lrDy, stKin.lrVeloY, stKin.lrAccelY));

END_FUNCTION

// ---- Test/FB_TravelTime_Test.TcPOU
// Tests for the travel-time formula behind the FEM 9.851 calculation.
FUNCTION_BLOCK FB_TravelTime_Test EXTENDS TcUnit.FB_TestSuite
VAR
    nDummy : INT;
END_VAR

Trapezoid_WhenTopSpeedIsReached();
Triangle_WhenTopSpeedIsNotReached();
NoDistance_TakesNoTime();

METHOD PRIVATE Trapezoid_WhenTopSpeedIsReached
VAR_INST
    bRan : BOOL;
END_VAR
TEST('Trapezoid_WhenTopSpeedIsReached');
IF bRan THEN
    TEST_FINISHED();
    RETURN;
END_IF
bRan := TRUE;

AssertEquals_LREAL(Expected := 20.0 / 3.0 + 3.0 / 0.6, Actual := F_TravelTime(20.0, 3.0, 0.6), Delta := 1.0E-9, Message := 's/v + v/a');

TEST_FINISHED();
END_METHOD

METHOD PRIVATE Triangle_WhenTopSpeedIsNotReached
VAR_INST
    bRan : BOOL;
END_VAR
TEST('Triangle_WhenTopSpeedIsNotReached');
IF bRan THEN
    TEST_FINISHED();
    RETURN;
END_IF
bRan := TRUE;

AssertEquals_LREAL(Expected := 2.0 * SQRT(1.0 / 0.6), Actual := F_TravelTime(1.0, 3.0, 0.6), Delta := 1.0E-9, Message := '2 * sqrt(s/a)');

TEST_FINISHED();
END_METHOD

METHOD PRIVATE NoDistance_TakesNoTime
VAR_INST
    bRan : BOOL;
END_VAR
TEST('NoDistance_TakesNoTime');
IF bRan THEN
    TEST_FINISHED();
    RETURN;
END_IF
bRan := TRUE;

AssertEquals_LREAL(Expected := 0.0, Actual := F_TravelTime(0.0, 3.0, 0.6), Delta := 1.0E-9, Message := 'zero distance');

TEST_FINISHED();
END_METHOD

END_FUNCTION_BLOCK

// ---- Test/FB_AxisNc_Test.TcPOU
// Tests for the NC axis path: FB_AxisNc on its own, and a whole RBG job with
// eAxisKind = eNc. They run against NC simulation axes (TestAxis, TestTravel,
// TestHoist, TestFork in the NC task), so unlike the other suites they take
// real time: one Cyclic() per PLC cycle until done or the cycle budget is spent.
FUNCTION_BLOCK FB_AxisNc_Test EXTENDS TcUnit.FB_TestSuite
VAR
    fbAxis   : FB_AxisNc(ipParent := 0, sNodeName := 'TestAxis');
    fbRackNc : FB_Rack;
    fbSrmNc  : FB_Srm(ipParent := 0, sNodeName := 'SrmNc');
END_VAR

MoveAbs_ReachesTheTargetOnTheNcAxis();
StoreJob_RunsOnNcAxes();

METHOD PRIVATE MoveAbs_ReachesTheTargetOnTheNcAxis
VAR_INST
    nCycles : DINT;
    eResult : E_CmdResult;
END_VAR
TEST('MoveAbs_ReachesTheTargetOnTheNcAxis');
fbAxis.bEnable    := TRUE;
fbAxis.lrVelocity := 1.0;
fbAxis.lrAccel    := 2.0;
eResult := fbAxis.MoveAbs(0.5);
fbAxis.Cyclic();
nCycles := nCycles + 1;
IF eResult = E_CmdResult.eBusy AND nCycles < 1000 THEN   // 10 s budget at 10 ms
    RETURN;
END_IF
AssertEquals_INT(Expected := TO_INT(E_CmdResult.eDone), Actual := TO_INT(eResult), Message := 'move must finish without error');
AssertEquals_LREAL(Expected := 0.5, Actual := fbAxis.ActPos, Delta := 0.002, Message := 'NC axis must stand at the target');
AssertFalse(Condition := fbAxis.Error, Message := 'no NC error');
TEST_FINISHED();
END_METHOD

METHOD PRIVATE StoreJob_RunsOnNcAxes
VAR_INST
    bStarted : BOOL;
    nCycles  : DINT;
END_VAR
VAR
    stStation : ST_SlotAddr := (nSide := 1, nColumn := 0, nLevel := 1);
    stPlace   : ST_SlotAddr := (nSide := 1, nColumn := 1, nLevel := 1);
END_VAR
TEST('StoreJob_RunsOnNcAxes');
IF NOT bStarted THEN
    bStarted := TRUE;
    fbSrmNc.eAxisKind := E_AxisKind.eNc;
    fbSrmNc.Init(fbRackNc);
    fbSrmNc.SetMode(E_OpMode.eAutomatic);
    fbRackNc.Put(stStation, 'LE0042');
    AssertTrue(Condition := fbSrmNc.StartJob(stStation, stPlace), Message := 'job must be accepted');
END_IF
fbSrmNc.Cyclic();
nCycles := nCycles + 1;
IF NOT fbSrmNc.bJobDone AND NOT fbSrmNc.bFault AND nCycles < 6000 THEN   // 60 s budget
    RETURN;
END_IF
AssertTrue(Condition := fbSrmNc.bJobDone, Message := 'store job on NC axes must finish');
AssertFalse(Condition := fbSrmNc.bFault, Message := 'no axis fault');
AssertEquals_STRING(Expected := 'LE0042', Actual := fbRackNc.LeIdAt(stPlace), Message := 'pallet must be booked into the place');
AssertEquals_LREAL(Expected := fbRackNc.TargetX(stPlace), Actual := fbSrmNc.TravelPos, Delta := 0.002, Message := 'RBG must stand at the place');
TEST_FINISHED();
END_METHOD

END_FUNCTION_BLOCK

// ---- Test/FB_HrlConfig_Test.TcPOU
// Tests for the plant configuration: parsing, range checks, defaults, and a
// rack of a different size built from the configuration without code changes.
FUNCTION_BLOCK FB_HrlConfig_Test EXTENDS TcUnit.FB_TestSuite
VAR
    fbCfgOk    : FB_HrlConfig;
    fbCfgBad   : FB_HrlConfig;
    fbCfgEmpty : FB_HrlConfig;
    fbCfgJunk  : FB_HrlConfig;
    fbSmallRack : FB_Rack;
END_VAR

Parse_ValidJson_SetsEveryGroup();
Parse_OutOfRangeValue_IsRejectedAndKeepsDefaults();
Parse_EmptyObject_GivesThePracticePlant();
Parse_NotJson_IsRejected();
SmallRack_FromConfig_LimitsAddressesAndSearch();

METHOD PRIVATE Parse_ValidJson_SetsEveryGroup
VAR
    sJson : STRING(1000) := '{"rack":{"sides":1,"columns":10,"levels":4,"pitchX":1.2},"axes":{"kind":"nc","travel":{"velocity":2.5,"accel":0.5}},"conveyors":{"infeed":{"length":1.8,"simulate":false}},"mfr":{"ackTimeout":8}}';
END_VAR
TEST('Parse_ValidJson_SetsEveryGroup');
AssertTrue(Condition := fbCfgOk.Parse(sJson), Message := 'valid config must parse');
AssertEquals_INT(Expected := 1, Actual := fbCfgOk.stConfig.stRack.nSides, Message := 'sides');
AssertEquals_INT(Expected := 10, Actual := fbCfgOk.stConfig.stRack.nColumns, Message := 'columns');
AssertEquals_INT(Expected := 4, Actual := fbCfgOk.stConfig.stRack.nLevels, Message := 'levels');
AssertEquals_LREAL(Expected := 1.2, Actual := fbCfgOk.stConfig.stRack.lrPitchX, Delta := 1.0E-9, Message := 'pitchX');
AssertEquals_LREAL(Expected := GVL_Rack.cPitchY, Actual := fbCfgOk.stConfig.stRack.lrPitchY, Delta := 1.0E-9, Message := 'missing pitchY keeps the default');
AssertTrue(Condition := fbCfgOk.stConfig.eAxisKind = E_AxisKind.eNc, Message := 'axes.kind nc');
AssertEquals_LREAL(Expected := 2.5, Actual := fbCfgOk.stConfig.stTravel.lrVelocity, Delta := 1.0E-9, Message := 'travel velocity');
AssertEquals_LREAL(Expected := 1.5, Actual := fbCfgOk.stConfig.stHoist.lrVelocity, Delta := 1.0E-9, Message := 'hoist keeps the default');
AssertEquals_LREAL(Expected := 1.8, Actual := fbCfgOk.stConfig.stInfeed.lrLength, Delta := 1.0E-9, Message := 'infeed length');
AssertFalse(Condition := fbCfgOk.stConfig.stInfeed.bSimulate, Message := 'infeed on real inputs');
AssertEquals_LREAL(Expected := 2.4, Actual := fbCfgOk.stConfig.stOutfeed.lrLength, Delta := 1.0E-9, Message := 'outfeed keeps the default');
AssertEquals_LREAL(Expected := 8.0, Actual := fbCfgOk.stConfig.lrAckTimeout, Delta := 1.0E-9, Message := 'ack timeout');
TEST_FINISHED();
END_METHOD

METHOD PRIVATE Parse_OutOfRangeValue_IsRejectedAndKeepsDefaults
VAR
    sJson : STRING(255) := '{"rack":{"columns":99},"axes":{"travel":{"velocity":2.0}}}';
END_VAR
TEST('Parse_OutOfRangeValue_IsRejectedAndKeepsDefaults');
AssertFalse(Condition := fbCfgBad.Parse(sJson), Message := '99 columns exceeds cMaxColumns');
AssertTrue(Condition := fbCfgBad.bError, Message := 'bError set');
AssertEquals_STRING(Expected := 'rack.columns out of range', Actual := fbCfgBad.sError, Message := 'error names the value');
AssertEquals_INT(Expected := GVL_Rack.cColumns, Actual := fbCfgBad.stConfig.stRack.nColumns, Message := 'columns stay default');
AssertEquals_LREAL(Expected := 3.0, Actual := fbCfgBad.stConfig.stTravel.lrVelocity, Delta := 1.0E-9, Message := 'a bad file never half-applies');
TEST_FINISHED();
END_METHOD

METHOD PRIVATE Parse_EmptyObject_GivesThePracticePlant
VAR
    sJson : STRING(10) := '{}';
END_VAR
TEST('Parse_EmptyObject_GivesThePracticePlant');
AssertTrue(Condition := fbCfgEmpty.Parse(sJson), Message := 'empty object is valid');
AssertEquals_INT(Expected := GVL_Rack.cColumns, Actual := fbCfgEmpty.stConfig.stRack.nColumns, Message := 'default columns');
AssertTrue(Condition := fbCfgEmpty.stConfig.eAxisKind = E_AxisKind.eSim, Message := 'default axes are simulated');
AssertTrue(Condition := fbCfgEmpty.stConfig.stInfeed.bSimulate, Message := 'default conveyors are simulated');
TEST_FINISHED();
END_METHOD

METHOD PRIVATE Parse_NotJson_IsRejected
VAR
    sJson : STRING(40) := 'columns = 10';
END_VAR
TEST('Parse_NotJson_IsRejected');
AssertFalse(Condition := fbCfgJunk.Parse(sJson), Message := 'plain text is not a config');
AssertTrue(Condition := fbCfgJunk.bError, Message := 'bError set');
TEST_FINISHED();
END_METHOD

METHOD PRIVATE SmallRack_FromConfig_LimitsAddressesAndSearch
VAR
    stAddr : ST_SlotAddr;
    stFree : ST_SlotAddr;
    nCol, nLvl, nSide : INT;
    nPut : INT;
END_VAR
TEST('SmallRack_FromConfig_LimitsAddressesAndSearch');
fbSmallRack.stCfg.nSides   := 2;
fbSmallRack.stCfg.nColumns := 10;
fbSmallRack.stCfg.nLevels  := 4;
stAddr.nSide := 1; stAddr.nColumn := 10; stAddr.nLevel := 4;
AssertTrue(Condition := fbSmallRack.IsValid(stAddr), Message := 'last place of a 10x4 rack is valid');
stAddr.nColumn := 11;
AssertFalse(Condition := fbSmallRack.IsValid(stAddr), Message := 'column 11 does not exist');
stAddr.nColumn := 1; stAddr.nLevel := 5;
AssertFalse(Condition := fbSmallRack.IsValid(stAddr), Message := 'level 5 does not exist');
FOR nCol := 1 TO 10 DO
    FOR nLvl := 1 TO 4 DO
        FOR nSide := 1 TO 2 DO
            stAddr.nSide := nSide; stAddr.nColumn := nCol; stAddr.nLevel := nLvl;
            IF fbSmallRack.Put(stAddr, 'LE') THEN
                nPut := nPut + 1;
            END_IF
        END_FOR
    END_FOR
END_FOR
AssertEquals_INT(Expected := 80, Actual := nPut, Message := '2 x 10 x 4 places');
AssertFalse(Condition := fbSmallRack.FindFree(stFree), Message := 'full small rack has no free place');
TEST_FINISHED();
END_METHOD

END_FUNCTION_BLOCK

// ---- Test/FB_TelegramCodec_Test.TcPOU
// Tests for the MFR wire format and for FB_MfrInterface.Serve over a link.
FUNCTION_BLOCK FB_TelegramCodec_Test EXTENDS TcUnit.FB_TestSuite
VAR
    fbCodec  : FB_TelegramCodec;
    fbCodec2 : FB_TelegramCodec;
    fbRack   : FB_Rack;
    fbSrm    : FB_Srm(ipParent := 0, sNodeName := 'SrmServe');
    fbMfr    : FB_MfrInterface;
    fbLink   : FB_MfrLinkFake;
    fbRackB  : FB_Rack;
    fbSrmB   : FB_Srm(ipParent := 0, sNodeName := 'SrmBad');
    fbMfrB   : FB_MfrInterface;
    fbLinkB  : FB_MfrLinkFake;
END_VAR

Encode_DefaultLayout_GivesTheDocumentedText();
Decode_RoundTrip_GivesTheSameTelegram();
Decode_WrongLength_IsRefused();
Decode_LetterInNumberField_IsRefused();
CustomLayout_ChangesLengthAndStillRoundTrips();
Serve_ValidOrder_AnswersTackOverTheLink();
Serve_BadFrame_AnswersTerr45();

// A transport order station -> place 2/4/3.
METHOD PRIVATE Order : ST_Telegram
VAR_INPUT
    nSeq : UINT;
END_VAR
Order.sType := 'TORD';
Order.nSeq  := nSeq;
Order.nOrder := 1234;
Order.sLeId := 'LE0042';
Order.stSource.nSide := 1; Order.stSource.nColumn := 0; Order.stSource.nLevel := 1;
Order.stTarget.nSide := 2; Order.stTarget.nColumn := 4; Order.stTarget.nLevel := 3;
Order.nStatus := 0;
END_METHOD

METHOD PRIVATE Encode_DefaultLayout_GivesTheDocumentedText
VAR
    sTxt : STRING(255);
END_VAR
TEST('Encode_DefaultLayout_GivesTheDocumentedText');
sTxt := fbCodec.Encode(Order(7));
AssertEquals_INT(Expected := 52, Actual := LEN(sTxt), Message := 'default telegram is 52 characters');
AssertEquals_STRING(Expected := 'TORD0000700001234LE0042              100001200403000', Actual := sTxt, Message := 'field order and padding');
TEST_FINISHED();
END_METHOD

METHOD PRIVATE Decode_RoundTrip_GivesTheSameTelegram
VAR
    stIn, stOut : ST_Telegram;
END_VAR
TEST('Decode_RoundTrip_GivesTheSameTelegram');
stIn := Order(7);
AssertTrue(Condition := fbCodec.Decode(fbCodec.Encode(stIn), stOut), Message := 'own text must decode');
AssertEquals_STRING(Expected := 'TORD', Actual := stOut.sType, Message := 'type');
AssertEquals_UINT(Expected := 7, Actual := stOut.nSeq, Message := 'seq');
AssertEquals_DINT(Expected := 1234, Actual := stOut.nOrder, Message := 'order');
AssertEquals_STRING(Expected := 'LE0042', Actual := stOut.sLeId, Message := 'load unit without padding');
AssertEquals_INT(Expected := 4, Actual := stOut.stTarget.nColumn, Message := 'target column');
AssertEquals_INT(Expected := 3, Actual := stOut.stTarget.nLevel, Message := 'target level');
TEST_FINISHED();
END_METHOD

METHOD PRIVATE Decode_WrongLength_IsRefused
VAR
    stOut : ST_Telegram;
END_VAR
TEST('Decode_WrongLength_IsRefused');
AssertFalse(Condition := fbCodec.Decode('TORD0000700001234', stOut), Message := 'short frame');
TEST_FINISHED();
END_METHOD

METHOD PRIVATE Decode_LetterInNumberField_IsRefused
VAR
    stOut : ST_Telegram;
END_VAR
TEST('Decode_LetterInNumberField_IsRefused');
AssertFalse(Condition := fbCodec.Decode('TORD0000700001234LE0042              10000120X403000', stOut), Message := 'X in the target column');
TEST_FINISHED();
END_METHOD

METHOD PRIVATE CustomLayout_ChangesLengthAndStillRoundTrips
VAR
    stOut : ST_Telegram;
    sTxt : STRING(255);
END_VAR
TEST('CustomLayout_ChangesLengthAndStillRoundTrips');
fbCodec2.stLayout.nOrder := 6;
fbCodec2.stLayout.nLeId  := 10;
sTxt := fbCodec2.Encode(Order(9));
AssertEquals_INT(Expected := 40, Actual := LEN(sTxt), Message := '52 - 2 - 10');
AssertTrue(Condition := fbCodec2.Decode(sTxt, stOut), Message := 'decodes with the same layout');
AssertEquals_DINT(Expected := 1234, Actual := stOut.nOrder, Message := 'order');
AssertFalse(Condition := fbCodec.Decode(sTxt, stOut), Message := 'default layout refuses it');
TEST_FINISHED();
END_METHOD

METHOD PRIVATE Serve_ValidOrder_AnswersTackOverTheLink
VAR
    stStation : ST_SlotAddr := (nSide := 1, nColumn := 0, nLevel := 1);
END_VAR
TEST('Serve_ValidOrder_AnswersTackOverTheLink');
fbSrm.Init(fbRack);
fbSrm.SetMode(E_OpMode.eAutomatic);
fbMfr.Init(fbRack, fbSrm);
fbRack.Put(stStation, 'LE0042');
fbLink.Give(Order(1));
fbMfr.Serve(fbLink);
AssertEquals_INT(Expected := 1, Actual := fbLink.nSent, Message := 'one answer sent');
AssertEquals_STRING(Expected := 'TACK', Actual := fbLink.aSent[1].sType, Message := 'order accepted');
AssertEquals_DINT(Expected := 1234, Actual := fbLink.aSent[1].nOrder, Message := 'answer names the order');
TEST_FINISHED();
END_METHOD

METHOD PRIVATE Serve_BadFrame_AnswersTerr45
VAR
    stBad : ST_Telegram;
END_VAR
TEST('Serve_BadFrame_AnswersTerr45');
fbSrmB.Init(fbRackB);
fbMfrB.Init(fbRackB, fbSrmB);
stBad.sType := 'BAD';
fbLinkB.Give(stBad);
fbMfrB.Serve(fbLinkB);
AssertEquals_STRING(Expected := 'TERR', Actual := fbLinkB.aSent[1].sType, Message := 'error answer');
AssertEquals_INT(Expected := GVL_Mfr.cUnknownTelegram, Actual := fbLinkB.aSent[1].nStatus, Message := 'status 45');
fbLinkB.Give(Order(1));
fbMfrB.Serve(fbLinkB);
AssertEquals_INT(Expected := GVL_Mfr.cSlotEmpty, Actual := fbLinkB.aSent[2].nStatus, Message := 'a bad frame does not use up sequence number 1');
TEST_FINISHED();
END_METHOD

END_FUNCTION_BLOCK

// ---- Test/FB_MfrLinkFake.TcPOU
// Test double for I_MfrLink: hands out one prepared telegram and records
// everything the PLC sends.
FUNCTION_BLOCK FB_MfrLinkFake IMPLEMENTS I_MfrLink
VAR
    stNext   : ST_Telegram;
    bHasNext : BOOL;
    aSent    : ARRAY[1..8] OF ST_Telegram;
    nSent    : INT;
END_VAR

METHOD PUBLIC Give
VAR_INPUT
    stTel : ST_Telegram;
END_VAR
stNext   := stTel;
bHasNext := TRUE;
END_METHOD

METHOD PUBLIC Poll : BOOL
VAR_IN_OUT
    stIn : ST_Telegram;
END_VAR
IF bHasNext THEN
    stIn     := stNext;
    bHasNext := FALSE;
    Poll     := TRUE;
END_IF
END_METHOD

METHOD PUBLIC Send : BOOL
VAR_INPUT
    stOut : ST_Telegram;
END_VAR
IF nSent < 8 THEN
    nSent := nSent + 1;
    aSent[nSent] := stOut;
    Send := TRUE;
END_IF
END_METHOD

PROPERTY PUBLIC Connected : BOOL
GET
Connected := TRUE;
END_GET
END_PROPERTY

END_FUNCTION_BLOCK

// ---- Test/FB_Operation_Test.TcPOU
// Tests for operation and commissioning: manual jog with interlock, guided
// teach-in, stop and resume of a job, and the fault list. Simulated axes,
// simulated time (whole scenario inside one PLC cycle).
FUNCTION_BLOCK FB_Operation_Test EXTENDS TcUnit.FB_TestSuite
VAR
    fbRackJog : FB_Rack;
    fbSrmJog  : FB_Srm(ipParent := 0, sNodeName := 'SrmJog');
    fbRackLock : FB_Rack;
    fbSrmLock  : FB_Srm(ipParent := 0, sNodeName := 'SrmLock');
    fbRackTeach : FB_Rack;
    fbSrmTeach  : FB_Srm(ipParent := 0, sNodeName := 'SrmTeach');
    fbTeach     : FB_TeachIn;
    fbRackStop : FB_Rack;
    fbSrmStop  : FB_Srm(ipParent := 0, sNodeName := 'SrmStop');
    fbDiag : FB_Diag;
END_VAR

Jog_Travel_MovesWhileHeldAndStopsOnRelease();
Jog_TravelWithForkOut_IsBlocked();
TeachIn_AtNominal_IsStoredAndFarOff_IsRefused();
Stop_DuringJob_HaltsAndAutomaticResumes();
Diag_FaultIsRaisedOncePerEdge();

METHOD PRIVATE Jog_Travel_MovesWhileHeldAndStopsOnRelease
VAR
    n : INT;
    lrHeld : LREAL;
END_VAR
TEST('Jog_Travel_MovesWhileHeldAndStopsOnRelease');
fbSrmJog.Init(fbRackJog);
fbSrmJog.SetMode(E_OpMode.eManual);
fbSrmJog.eJogAxis := E_JogAxis.eTravel;
fbSrmJog.bJogFwd  := TRUE;
FOR n := 1 TO 200 DO      // 2 s simulated
    fbSrmJog.Cyclic();
END_FOR
lrHeld := fbSrmJog.TravelPos;
AssertTrue(Condition := lrHeld > 0.5, Message := 'travel moves while the button is held');
fbSrmJog.bJogFwd := FALSE;
FOR n := 1 TO 200 DO
    fbSrmJog.Cyclic();
END_FOR
AssertEquals_LREAL(Expected := lrHeld, Actual := fbSrmJog.TravelPos, Delta := 0.05, Message := 'travel stops on release');
TEST_FINISHED();
END_METHOD

METHOD PRIVATE Jog_TravelWithForkOut_IsBlocked
VAR
    n : INT;
END_VAR
TEST('Jog_TravelWithForkOut_IsBlocked');
fbSrmLock.Init(fbRackLock);
fbSrmLock.SetMode(E_OpMode.eManual);
fbSrmLock.eJogAxis := E_JogAxis.eFork;
fbSrmLock.bJogFwd  := TRUE;
FOR n := 1 TO 100 DO      // fork out by about 0.3 m
    fbSrmLock.Cyclic();
END_FOR
fbSrmLock.bJogFwd := FALSE;
fbSrmLock.Cyclic();
AssertTrue(Condition := fbSrmLock.ForkActPos > 0.1, Message := 'fork is out');
fbSrmLock.eJogAxis := E_JogAxis.eTravel;
fbSrmLock.bJogFwd  := TRUE;
FOR n := 1 TO 100 DO
    fbSrmLock.Cyclic();
END_FOR
AssertTrue(Condition := fbSrmLock.bJogBlocked, Message := 'interlock reported');
AssertEquals_LREAL(Expected := 0.0, Actual := fbSrmLock.TravelPos, Delta := 0.001, Message := 'travel must not move with the fork out');
TEST_FINISHED();
END_METHOD

METHOD PRIVATE TeachIn_AtNominal_IsStoredAndFarOff_IsRefused
VAR
    stPlace : ST_SlotAddr := (nSide := 1, nColumn := 2, nLevel := 2);
    stFar   : ST_SlotAddr := (nSide := 1, nColumn := 3, nLevel := 2);
    n : INT;
END_VAR
TEST('TeachIn_AtNominal_IsStoredAndFarOff_IsRefused');
fbSrmTeach.Init(fbRackTeach);
fbSrmTeach.SetMode(E_OpMode.eManual);
fbTeach.Init(fbRackTeach, fbSrmTeach);
AssertTrue(Condition := fbTeach.Start(stPlace), Message := 'teach start accepted');
FOR n := 1 TO 3000 DO
    fbSrmTeach.Cyclic();
    IF NOT fbSrmTeach.bGotoActive THEN EXIT; END_IF
END_FOR
AssertEquals_LREAL(Expected := fbRackTeach.NominalX(stPlace), Actual := fbSrmTeach.TravelPos, Delta := 0.002, Message := 'RBG at the nominal place');
AssertTrue(Condition := fbTeach.Confirm(), Message := 'position within tolerance is stored');
AssertEquals_INT(Expected := 1, Actual := fbTeach.nTaught, Message := 'one place taught');
// Next place: drive there, then the operator jogs the hoist about 0.1 m too high.
fbTeach.Start(stFar);
AssertFalse(Condition := fbTeach.Confirm(), Message := 'still driving: no confirm');
FOR n := 1 TO 3000 DO
    fbSrmTeach.Cyclic();
    IF NOT fbSrmTeach.bGotoActive THEN EXIT; END_IF
END_FOR
fbSrmTeach.eJogAxis := E_JogAxis.eHoist;
fbSrmTeach.bJogFwd  := TRUE;
FOR n := 1 TO 50 DO
    fbSrmTeach.Cyclic();
END_FOR
fbSrmTeach.bJogFwd := FALSE;
fbSrmTeach.Cyclic();
AssertFalse(Condition := fbTeach.Confirm(), Message := 'far from the drawing: refused');
AssertTrue(Condition := fbTeach.bLastRejected, Message := 'rejection reported');
TEST_FINISHED();
END_METHOD

METHOD PRIVATE Stop_DuringJob_HaltsAndAutomaticResumes
VAR
    stStation : ST_SlotAddr := (nSide := 1, nColumn := 0, nLevel := 1);
    stPlace   : ST_SlotAddr := (nSide := 2, nColumn := 6, nLevel := 3);
    n : DINT;
    lrStopped : LREAL;
END_VAR
TEST('Stop_DuringJob_HaltsAndAutomaticResumes');
fbSrmStop.Init(fbRackStop);
fbSrmStop.SetMode(E_OpMode.eAutomatic);
fbRackStop.Put(stStation, 'LE0007');
fbSrmStop.StartJob(stStation, stPlace);
FOR n := 1 TO 300 DO
    fbSrmStop.Cyclic();
END_FOR
fbSrmStop.SetMode(E_OpMode.eStop);
fbSrmStop.Cyclic();
lrStopped := fbSrmStop.TravelPos;
FOR n := 1 TO 300 DO
    fbSrmStop.Cyclic();
END_FOR
AssertEquals_LREAL(Expected := lrStopped, Actual := fbSrmStop.TravelPos, Delta := 0.001, Message := 'no motion in stop');
AssertTrue(Condition := fbSrmStop.bBusy, Message := 'job still pending');
fbSrmStop.SetMode(E_OpMode.eAutomatic);
FOR n := 1 TO 30000 DO
    fbSrmStop.Cyclic();
    IF fbSrmStop.bJobDone OR fbSrmStop.bFault THEN EXIT; END_IF
END_FOR
AssertEquals_STRING(Expected := 'LE0007', Actual := fbRackStop.LeIdAt(stPlace), Message := 'job finishes after automatic again');
TEST_FINISHED();
END_METHOD

METHOD PRIVATE Diag_FaultIsRaisedOncePerEdge
VAR
END_VAR
TEST('Diag_FaultIsRaisedOncePerEdge');
fbDiag.Check(E_Fault.eInfeedJam, TRUE, 'test jam');
fbDiag.Check(E_Fault.eInfeedJam, TRUE, 'test jam');
AssertEquals_UDINT(Expected := 1, Actual := fbDiag.nRaised, Message := 'raised once while active');
AssertEquals_INT(Expected := 1, Actual := fbDiag.nActive, Message := 'one active');
AssertEquals_STRING(Expected := 'test jam', Actual := fbDiag.aText[TO_INT(E_Fault.eInfeedJam)], Message := 'text for the HMI');
fbDiag.Check(E_Fault.eInfeedJam, FALSE, 'test jam');
AssertEquals_INT(Expected := 0, Actual := fbDiag.nActive, Message := 'cleared');
AssertEquals_STRING(Expected := '', Actual := fbDiag.aText[TO_INT(E_Fault.eInfeedJam)], Message := 'text cleared');
TEST_FINISHED();
END_METHOD

END_FUNCTION_BLOCK

// ---- Test/FB_SafetyInterface_Test.TcPOU
// Tests for the standard-PLC side of the safety concept (not the safety
// function itself): every drop disables, no restart without acknowledge,
// door unlock only at standstill.
FUNCTION_BLOCK FB_SafetyInterface_Test EXTENDS TcUnit.FB_TestSuite
VAR
    fbStart : FB_SafetyInterface;
    fbDrop  : FB_SafetyInterface;
    fbDoor  : FB_SafetyInterface;
END_VAR

PowerUp_NeedsAcknowledgeBeforeEnable();
EveryDrop_DisablesAndLocksUntilReset();
DoorUnlock_OnlyAtStandstill();

METHOD PRIVATE AllOk : ST_SafetyStatus
VAR_INPUT
END_VAR
AllOk.bSafetyRun  := TRUE;
AllOk.bEStopOk    := TRUE;
AllOk.bDoorClosed := TRUE;
AllOk.bDoorLocked := TRUE;
AllOk.bStoOk      := TRUE;
END_METHOD

METHOD PRIVATE PowerUp_NeedsAcknowledgeBeforeEnable
VAR
END_VAR
TEST('PowerUp_NeedsAcknowledgeBeforeEnable');
fbStart(stStatus := AllOk(), bReset := FALSE);
AssertFalse(Condition := fbStart.bDriveEnable, Message := 'no enable straight after power-up');
fbStart(stStatus := AllOk(), bReset := TRUE);
AssertTrue(Condition := fbStart.bDriveEnable, Message := 'enable after acknowledge');
TEST_FINISHED();
END_METHOD

METHOD PRIVATE EveryDrop_DisablesAndLocksUntilReset
VAR
    stSt : ST_SafetyStatus;
    i : INT;
END_VAR
TEST('EveryDrop_DisablesAndLocksUntilReset');
fbDrop(stStatus := AllOk(), bReset := TRUE);   // running
fbDrop(stStatus := AllOk(), bReset := FALSE);
FOR i := 1 TO 5 DO
    stSt := AllOk();
    CASE i OF
        1: stSt.bSafetyRun  := FALSE;
        2: stSt.bEStopOk    := FALSE;
        3: stSt.bDoorClosed := FALSE;
        4: stSt.bDoorLocked := FALSE;
        5: stSt.bStoOk      := FALSE;
    END_CASE
    fbDrop(stStatus := stSt, bReset := FALSE);
    AssertFalse(Condition := fbDrop.bDriveEnable, Message := 'a dropped bit disables');
    fbDrop(stStatus := AllOk(), bReset := FALSE);
    AssertFalse(Condition := fbDrop.bDriveEnable, Message := 'bit back: still locked, no automatic restart');
    AssertTrue(Condition := fbDrop.bRestartLock, Message := 'restart lock set');
    fbDrop(stStatus := stSt, bReset := TRUE);
    AssertFalse(Condition := fbDrop.bDriveEnable, Message := 'reset while still dropped does nothing');
    fbDrop(stStatus := AllOk(), bReset := FALSE);
    fbDrop(stStatus := AllOk(), bReset := TRUE);
    AssertTrue(Condition := fbDrop.bDriveEnable, Message := 'reset with all OK enables');
    fbDrop(stStatus := AllOk(), bReset := FALSE);
END_FOR
TEST_FINISHED();
END_METHOD

METHOD PRIVATE DoorUnlock_OnlyAtStandstill
VAR
END_VAR
TEST('DoorUnlock_OnlyAtStandstill');
fbDoor(stStatus := AllOk(), bDoorRequest := TRUE, bStandstill := FALSE);
AssertFalse(Condition := fbDoor.bDoorUnlockReq, Message := 'no unlock while the RBG moves');
fbDoor(stStatus := AllOk(), bDoorRequest := TRUE, bStandstill := TRUE);
AssertTrue(Condition := fbDoor.bDoorUnlockReq, Message := 'unlock request at standstill');
TEST_FINISHED();
END_METHOD

END_FUNCTION_BLOCK
